(* IEC 61131-3 sources: iecf/harness/cases (part 5) *)

(* ---- narrowingcompare.st ---- *)
(* implicit-narrowing: a ULINT and a signed integer, which no type holds
   both of, compared by their values, W0010 at each - as TcOpen's tests'
   `_plcCycleCounter >= _reqStep + 7`, a ULINT and an INT. Worked by
   hand, u 5, m -1, big 2^64 - 1, l -1, seven 7, four 4:
   u > m TRUE (%QX0.0); m < u TRUE (%QX0.1); u = m FALSE (%QX0.2);
   big > l TRUE, where the bits alike would say equal (%QX0.3);
   u + 2 = seven, 7 = 7, TRUE (%QX0.4); u <= four FALSE (%QX0.5).
   reference-skip: implicit narrowing is CODESYS's, not IEC 61131-3. *)
PROGRAM main
  VAR
    u : ULINT := 5; big : ULINT := 18446744073709551615;
    m : INT := -1; l : LINT := -1; seven : DINT := 7; four : SINT := 4;
  END_VAR
  VAR
    q0 AT %QX0.0 : BOOL; q1 AT %QX0.1 : BOOL; q2 AT %QX0.2 : BOOL;
    q3 AT %QX0.3 : BOOL; q4 AT %QX0.4 : BOOL; q5 AT %QX0.5 : BOOL;
  END_VAR
  q0 := u > m;
  q1 := m < u;
  q2 := u = m;
  q3 := big > l;
  q4 := u + 2 = seven;
  q5 := u <= four;
END_PROGRAM

CONFIGURATION cf
  RESOURCE r ON x
    TASK tk(INTERVAL := T#10ms, PRIORITY := 1);
    PROGRAM p WITH tk : main;
  END_RESOURCE
END_CONFIGURATION

(* ---- narrowingliteral.st ---- *)
(* implicit-narrowing: an integer literal outside the integer or bit
   string type it goes into keeps its low bits, as a conversion of a
   typed one would, W0010 at each - as TcOpen's `_testId := -1` of a
   ULINT and `_theOrderOfThePreviouslyExecutedStep := -1` of a UINT.
   Worked by hand:
   u := -1, a UINT: 65535, 16#FFFF (%QW0).
   g(300), to a USINT input: 300 - 256, 44, 16#2C (%QB2).
   s := 200, a SINT: 200 - 256, -56, 16#C8 (%QB3).
   w := 16#12345, a WORD: 16#2345 (%QW4).
   l := -1, a ULINT: 2^64 - 1, all ones (%QL8).
   i, initialised to -2, a UDINT: 2^32 - 2, 16#FFFFFFFE (%QD16).
   reference-skip: implicit narrowing is CODESYS's, not IEC 61131-3. *)
FUNCTION g : USINT
  VAR_INPUT x : USINT; END_VAR
  g := x;
END_FUNCTION

PROGRAM main
  VAR
    u : UINT; s : SINT; w : WORD; l : ULINT; i : UDINT := -2;
  END_VAR
  VAR
    q0 AT %QW0 : UINT; q1 AT %QB2 : USINT; q2 AT %QB3 : SINT; q3 AT %QW4 : WORD;
    q4 AT %QL8 : ULINT; q5 AT %QD16 : UDINT;
  END_VAR
  u := -1;
  q0 := u;
  q1 := g(300);
  s := 200;
  q2 := s;
  w := 16#12345;
  q3 := w;
  l := -1;
  q4 := l;
  q5 := i;
END_PROGRAM

CONFIGURATION cf
  RESOURCE r ON x
    TASK tk(INTERVAL := T#10ms, PRIORITY := 1);
    PROGRAM p WITH tk : main;
  END_RESOURCE
END_CONFIGURATION

(* ---- narrowingreal.st ---- *)
(* implicit-narrowing: an integer where a real is wanted and Figure 11
   has no implicit conversion, and an LREAL where a REAL is, converted
   as DINT_TO_REAL and LREAL_TO_REAL would, W0010 at each - as TcOpen's
   `_price := Price` (an LREAL property into a REAL), its
   TcoBytesToReal's LREAL into the REAL result, and a DINT given to
   TcoRealToBytes's `inValue : REAL`. Worked by hand:
   r := d, DINT 16777217 into a REAL: the nearest REAL, 16777216.0,
   16#4B800000 (%QD0).
   r := l, LREAL 1.5: 1.5, 16#3FC00000 (%QD4).
   twice(n), the DINT 3 to a REAL input: 6.0, 16#40C00000 (%QD8).
   quarter(), an LREAL 2.25 into the REAL result: 16#40100000 (%QD12).
   reference-skip: implicit narrowing is CODESYS's, not IEC 61131-3. *)
FUNCTION twice : REAL
  VAR_INPUT x : REAL; END_VAR
  twice := x * 2.0;
END_FUNCTION

FUNCTION quarter : REAL
  VAR l : LREAL := 2.25; END_VAR
  quarter := l;
END_FUNCTION

PROGRAM main
  VAR
    d : DINT := 16777217; l : LREAL := 1.5; n : DINT := 3; r : REAL;
  END_VAR
  VAR
    q0 AT %QD0 : REAL;
    q1 AT %QD4 : REAL;
    q2 AT %QD8 : REAL;
    q3 AT %QD12 : REAL;
  END_VAR
  r := d;
  q0 := r;
  r := l;
  q1 := r;
  q2 := twice(n);
  q3 := quarter();
END_PROGRAM

CONFIGURATION cf
  RESOURCE r ON x
    TASK tk(INTERVAL := T#10ms, PRIORITY := 1);
    PROGRAM p WITH tk : main;
  END_RESOURCE
END_CONFIGURATION

(* ---- nesten.st ---- *)
(* Calls with EN nested in another's arguments, and EN on a FUNCTION
   giving an array or a structure (Ed.3 6.6.1.5; docs/dependencies.md:
   EN FALSE does not evaluate the inputs, calls nothing and leaves the
   statement undone). Worked by hand:
   b TRUE: ADD(EN := b, IN1 := ADD(EN := b, IN1 := 1, IN2 := 2),
   IN2 := 3): 6 (%QB0). b FALSE, v 9 before: the statement is undone, v
   9 (%QB1).
   t 32767: ADD(EN := TRUE, IN1 := ADD(EN := TRUE, IN1 := t, IN2 := 1,
   ENO => e2), IN2 := 0, ENO => e1): the inner one overflows, wraps to
   -32768 and is flagged OVERFLOW, its ENO FALSE (%QX2.0 0); the outer
   adds 0, no flag of its own: its ENO TRUE (%QX2.1 1); v / 1000 is -32
   (%QB3).
   Inc adds 1 to its in-out. n 0: ADD(EN := TRUE, IN1 := Inc(EN :=
   TRUE, io := n), IN2 := 10): 11 (%QB4), n 1 (%QB5). The outer's EN
   FALSE, v 5 before: Inc is not called, v 5 (%QB6), n still 1 (%QB7).
   FA gives [x, 2x, 0]: a := FA(EN := TRUE, x := 4), a[2] 8 (%QB8);
   a := FA(EN := FALSE, x := 7) leaves a: a[1] 4 (%QB9).
   p := FP(EN := TRUE, x := 3, ENO => e3): p.x 3 (%QB10), e3 TRUE
   (%QX11.0). SumA(FA(EN := TRUE, x := 2)), 2 + 4 + 0: 6 (%QB12).
   The first flag is the inner ADD's OVERFLOW.
   reference-skip: a nested call with ENO or an in-out, an array
   input: its C does not build. *)
TYPE
  A3 : ARRAY [1..3] OF INT;
  PT : STRUCT x : INT; END_STRUCT;
END_TYPE
FUNCTION Inc : INT
  VAR_IN_OUT io : INT; END_VAR
  io := io + 1;
  Inc := io;
END_FUNCTION
FUNCTION FA : A3
  VAR_INPUT x : INT; END_VAR
  FA[1] := x;
  FA[2] := x * 2;
END_FUNCTION
FUNCTION FP : PT
  VAR_INPUT x : INT; END_VAR
  FP.x := x;
END_FUNCTION
FUNCTION SumA : INT
  VAR_INPUT q : A3; END_VAR
  SumA := q[1] + q[2] + q[3];
END_FUNCTION
PROGRAM main
  VAR
    b : BOOL := TRUE;
    v : INT;
    t : INT := 32767;
    n : INT;
    e1 : BOOL;
    e2 : BOOL;
    e3 : BOOL;
    a : A3;
    p : PT;
  END_VAR
  VAR
    q0 AT %QB0 : SINT;
    q1 AT %QB1 : SINT;
    q20 AT %QX2.0 : BOOL;
    q21 AT %QX2.1 : BOOL;
    q3 AT %QB3 : SINT;
    q4 AT %QB4 : SINT;
    q5 AT %QB5 : SINT;
    q6 AT %QB6 : SINT;
    q7 AT %QB7 : SINT;
    q8 AT %QB8 : SINT;
    q9 AT %QB9 : SINT;
    q10 AT %QB10 : SINT;
    q11 AT %QX11.0 : BOOL;
    q12 AT %QB12 : SINT;
  END_VAR
  v := ADD(EN := b, IN1 := ADD(EN := b, IN1 := 1, IN2 := 2), IN2 := 3);
  q0 := INT_TO_SINT(v);
  b := FALSE;
  v := 9;
  v := ADD(EN := b, IN1 := ADD(EN := b, IN1 := 1, IN2 := 2), IN2 := 3);
  q1 := INT_TO_SINT(v);
  v := ADD(EN := TRUE, IN1 := ADD(EN := TRUE, IN1 := t, IN2 := 1, ENO => e2), IN2 := 0, ENO => e1);
  q20 := e2;
  q21 := e1;
  q3 := INT_TO_SINT(v / 1000);
  n := 0;
  v := ADD(EN := TRUE, IN1 := Inc(EN := TRUE, io := n), IN2 := 10);
  q4 := INT_TO_SINT(v);
  q5 := INT_TO_SINT(n);
  v := 5;
  v := ADD(EN := FALSE, IN1 := Inc(EN := TRUE, io := n), IN2 := 10);
  q6 := INT_TO_SINT(v);
  q7 := INT_TO_SINT(n);
  a := FA(EN := TRUE, x := 4);
  q8 := INT_TO_SINT(a[2]);
  a := FA(EN := FALSE, x := 7);
  q9 := INT_TO_SINT(a[1]);
  p := FP(EN := TRUE, x := 3, ENO => e3);
  q10 := INT_TO_SINT(p.x);
  q11 := e3;
  q12 := INT_TO_SINT(SumA(FA(EN := TRUE, x := 2)));
END_PROGRAM

CONFIGURATION c
  RESOURCE r ON x
    TASK t(INTERVAL := T#10ms, PRIORITY := 1);
    PROGRAM p WITH t : main;
  END_RESOURCE
END_CONFIGURATION

(* ---- overflow.st ---- *)
(* Where iecf differs from the reference compiler on purpose (PROPOSAL.md §6.3): an
   integer overflow is flagged. At tick 2, a + b leaves INT. Both wrap to
   -1536 and go on, as CODESYS, TwinCAT, Siemens and Rockwell do; iecf
   also records the first overflow, its POU and line, in ctx->flag, which
   stays until the platform clears it. Its trace is overflow.iecf.trace:
   the reference compiler's bytes, with "flag 2 MAIN 18" from tick 2.

   MOD by zero is 0 in both: Ed.3 Table 29 e defines it so. *)
PROGRAM main
VAR
  a AT %IW0 : INT;
  b AT %IW2 : INT;
  r_mod AT %MW0 : INT;
  r_sum AT %MW2 : INT;
  after AT %MW4 : INT;
END_VAR
r_mod := a MOD b;
r_sum := a + b;
after := after + 1;
END_PROGRAM

CONFIGURATION plant
  RESOURCE r ON PLC
    TASK fast(INTERVAL := T#10ms, PRIORITY := 0);
    PROGRAM p WITH fast : main;
  END_RESOURCE
END_CONFIGURATION

(* ---- parts.st ---- *)
(* CONCAT_DATE, CONCAT_TOD, CONCAT_DT and the SPLITs (Ed.3 Table 36;
   docs/dependencies.md): a month from 11 and an hour from 22 go up by one
   each tick, joined into a DATE, a TOD and a DT and split back. The parts
   are valid at tick 1 (2026-12-31, 23:30:15.250); a day not in its month
   (November 31st, at tick 0), a month 13 or an hour 24 gives the type's
   default value in iecf, flagged; iecf's trace is parts.iecf.trace. *)
PROGRAM main
VAR
  r_year AT %MW0 : UINT;
  r_month AT %MB2 : USINT;
  r_day AT %MB3 : USINT;
  r_hour AT %MB4 : USINT;
  r_min AT %MB5 : USINT;
  r_sec AT %MB6 : USINT;
  r_ms AT %MW8 : UINT;
  r_dt_month AT %MB10 : USINT;
  r_dt_hour AT %MB11 : USINT;
END_VAR
VAR
  month : INT := 10;
  hour : SINT := 21;
  d : DATE;
  t : TOD;
  s : DT;
  y, m, dd : UDINT;
END_VAR
month := month + 1;
hour := hour + 1;
d := CONCAT_DATE(2026, month, 31);
t := CONCAT_TOD(hour, 30, 15, 250);
s := CONCAT_DT(YEAR := 2026, MONTH := month, DAY := 28, HOUR := hour,
               MINUTE := 59, SECOND := 59, MILLISECOND := 999);
SPLIT_DATE(d, y, m, dd);
r_year := UDINT_TO_UINT(y);
r_month := UDINT_TO_USINT(m);
r_day := UDINT_TO_USINT(dd);
SPLIT_TOD(IN := t, HOUR => r_hour, MINUTE => r_min, SECOND => r_sec, MILLISECOND => r_ms);
SPLIT_DT(IN := s, MONTH => r_dt_month, HOUR => r_dt_hour);
END_PROGRAM

CONFIGURATION plant
  RESOURCE r ON PLC
    TASK fast(INTERVAL := T#10ms, PRIORITY := 0);
    PROGRAM p WITH fast : main;
  END_RESOURCE
END_CONFIGURATION

(* ---- pointerfault.st ---- *)
(* A pointer read past its variable (the pointers extension): a fault,
   IECF_FAULT_INDEX, the task stopped where the read leaves the variable,
   never C's undefined behaviour. Worked by hand: a has 4 bytes, 1 2 3 4;
   the loop adds them through pt for i 0..4, so the fifth read, past the
   end, faults on line 21 in the first tick, n holding 10 so far, and
   the task stops there: %QB0, set after the loop, stays 0. (The host
   leaves the fault set, so a later tick stops at once: whether to run
   again is the platform's; %QB1 is the first statement's, 0.)
   reference-skip: pointers are CODESYS's, not IEC 61131-3. *)
PROGRAM main
  VAR
    a : ARRAY[0..3] OF BYTE := [1, 2, 3, 4];
    pt : POINTER TO BYTE;
    i, n : INT;
  END_VAR
  VAR q0 AT %QB0 : SINT; q1 AT %QB1 : SINT; END_VAR
  q1 := INT_TO_SINT(n);
  n := 0;
  pt := ADR(a);
  FOR i := 0 TO 4 DO
    n := n + BYTE_TO_INT(pt^);
    pt := pt + 1;
  END_FOR;
  q0 := INT_TO_SINT(n);
END_PROGRAM

CONFIGURATION cf
  RESOURCE r ON x
    TASK tk(INTERVAL := T#10ms, PRIORITY := 1);
    PROGRAM p WITH tk : main;
  END_RESOURCE
END_CONFIGURATION

(* ---- pointerindex.st ---- *)
(* A pointer indexed (the pointers extension): p[i] is (p + i *
   SIZEOF(T))^, as CODESYS and TwinCAT index a pointer, checked as p^
   is. Worked by hand: a is 10 20 30 40 50, so the loop adds 150 and
   %QB0 is 15; p[k] with k 2 writes a[2] := 7; p moved to ADR(p[3]),
   a[3], reads p[-1] + p[0], 7 + 40, so %QB1 is 47; q[1].y := 9 and
   s[2].x := 4 read back through q and s, 9 + 4, %QB2 13; p[1] is
   a[4], 50, %QB3 5; %QB4 set to 1, then p[2] is past a's end: a
   fault, IECF_FAULT_INDEX, on line 36, %QB4 left at 1.
   reference-skip: pointers are CODESYS's, not IEC 61131-3. *)
TYPE pair : STRUCT x : INT; y : INT; END_STRUCT; END_TYPE
PROGRAM main
  VAR
    a : ARRAY[0..4] OF INT := [10, 20, 30, 40, 50];
    s : ARRAY[0..2] OF pair;
    p : POINTER TO INT;
    q : POINTER TO pair;
    i, n : INT;
    k : UINT := 2;
  END_VAR
  VAR q0 AT %QB0 : SINT; q1 AT %QB1 : SINT; q2 AT %QB2 : SINT; q3 AT %QB3 : SINT; q4 AT %QB4 : SINT; END_VAR
  p := ADR(a);
  n := 0;
  FOR i := 0 TO 4 DO
    n := n + p[i];
  END_FOR;
  q0 := INT_TO_SINT(n / 10);
  p[k] := 7;
  p := ADR(p[3]);
  q1 := INT_TO_SINT(p[-1] + p[0]);
  q := ADR(s);
  q[1].y := 9;
  s[2].x := 4;
  q2 := INT_TO_SINT(s[1].y + q[2].x);
  q3 := INT_TO_SINT(p[1] / 10);
  q4 := 1;
  q4 := INT_TO_SINT(p[2]);
END_PROGRAM

CONFIGURATION cf
  RESOURCE r ON x
    TASK tk(INTERVAL := T#10ms, PRIORITY := 1);
    PROGRAM p WITH tk : main;
  END_RESOURCE
END_CONFIGURATION

(* ---- pointers.st ---- *)
(* Pointers (the pointers extension), in the ways the OSCAT BASIC library
   uses them. Worked by hand:
   %QB0: StrLen walks a STRING's bytes through a POINTER TO BYTE to its
   0: 'hello', 5.
   %QB1: Sum takes ADR(a) and SIZEOF(a) of an ARRAY[0..3] OF REAL, as
   OSCAT's array functions do, and counts SIZEOF(a) / SIZEOF(pt^[0]) = 4
   elements: 1.5 + 2.5 + 3.0 + 4.0 = 11.0, as SINT 11.
   %QB2: Clear zeroes a BYTE buffer by pointer arithmetic, pt < stop,
   pt := pt + 1, from ADR(buf) to ADR(buf) + SIZEOF(buf); then buf[0] +
   buf[7], 0.
   %QB3: four bytes 16#11 16#22 16#33 16#44 read as one DWORD through a
   POINTER TO DWORD: 16#44332211 on a little-endian platform, its low
   byte 16#11.
   %QB4: a structure's field through a pointer, s.b := 7 by ps^.b := 7;
   and ps^.a + ps^.b with a 2: 9.
   %QB5: two pointers into one array subtracted: ADR(a[3]) - ADR(a[0]),
   3 * SIZEOF(REAL), 12.
   reference-skip: pointers are CODESYS's, not IEC 61131-3. *)
TYPE Pair : STRUCT a : SINT; b : SINT; END_STRUCT; END_TYPE

FUNCTION StrLen : INT
  VAR_INPUT pt : POINTER TO BYTE; END_VAR
  StrLen := 0;
  WHILE pt^ <> 0 DO
    StrLen := StrLen + 1;
    pt := pt + 1;
  END_WHILE;
END_FUNCTION

FUNCTION Sum : REAL
  VAR_INPUT pt : POINTER TO ARRAY[0..32000] OF REAL; size : UINT; END_VAR
  VAR i : INT; END_VAR
  Sum := 0.0;
  FOR i := 0 TO UINT_TO_INT(size / SIZEOF(pt^[0])) - 1 DO
    Sum := Sum + pt^[i];
  END_FOR;
END_FUNCTION

FUNCTION Clear : BOOL
  VAR_INPUT pt : POINTER TO BYTE; size : UINT; END_VAR
  VAR stop : POINTER TO BYTE; END_VAR
  stop := pt + size;
  WHILE pt < stop DO
    pt^ := 0;
    pt := pt + 1;
  END_WHILE;
  Clear := TRUE;
END_FUNCTION

PROGRAM main
  VAR
    s : STRING[20] := 'hello';
    a : ARRAY[0..3] OF REAL := [1.5, 2.5, 3.0, 4.0];
    buf : ARRAY[0..7] OF BYTE := [8(16#FF)];
    bytes : ARRAY[0..3] OF BYTE := [16#11, 16#22, 16#33, 16#44];
    pd : POINTER TO DWORD;
    pr : Pair := (a := 2);
    ps : POINTER TO Pair;
    ok : BOOL;
  END_VAR
  VAR
    q0 AT %QB0 : SINT; q1 AT %QB1 : SINT; q2 AT %QB2 : BYTE; q3 AT %QB3 : BYTE;
    q4 AT %QB4 : SINT; q5 AT %QB5 : SINT;
  END_VAR
  q0 := INT_TO_SINT(StrLen(ADR(s)));
  q1 := REAL_TO_SINT(Sum(ADR(a), SIZEOF(a)));
  ok := Clear(ADR(buf), SIZEOF(buf));
  q2 := buf[0] OR buf[7];
  pd := ADR(bytes);
  q3 := DWORD_TO_BYTE(pd^);
  ps := ADR(pr);
  ps^.b := 7;
  q4 := ps^.a + ps^.b;
  q5 := DINT_TO_SINT(ADR(a[3]) - ADR(a[0]));
END_PROGRAM

CONFIGURATION cf
  RESOURCE r ON x
    TASK tk(INTERVAL := T#10ms, PRIORITY := 1);
    PROGRAM p WITH tk : main;
  END_RESOURCE
END_CONFIGURATION

(* ---- pointers2.st ---- *)
(* Pointers (the pointers extension): a STRING whole through a pointer,
   arrays and structures copied whole through one, ADR of a variable at
   an address, and ADR() as an initial value. Worked by hand:
   %QB0: ps := ADR(s); ps^ := 'abc' writes the STRING through ps; then
   LEN(s), 3.
   %QB1: t := ps^ reads it back whole; LEN(t) + LEN(ps^), 3 + 3 = 6.
   %QB2: pa := ADR(src); dst := pa^ copies the array [5, 6, 7] whole;
   dst[2], 7.
   %QB3: pq^ := pr copies a structure whole into r2 (pq := ADR(r2)), then
   r2.b, 9.
   %QB4: pin points at %IB2, ADR of a variable at an address; the
   input bytes are 0, so pin^ reads 0; pq0 points at the output %QB5 and
   writes 16#2A through it (%QB5), read back as 42 into %QB4.
   %QB6: pinit's initial value ADR(src[1]) points at src[1], 6.
   reference-skip: pointers are CODESYS's, not IEC 61131-3. *)
TYPE R : STRUCT a : SINT; b : SINT; END_STRUCT; END_TYPE

PROGRAM main
  VAR
    s : STRING[20];
    t : STRING[20];
    ps : POINTER TO STRING[20];
    src : ARRAY[0..2] OF SINT := [5, 6, 7];
    dst : ARRAY[0..2] OF SINT;
    pa : POINTER TO ARRAY[0..2] OF SINT;
    pr : R := (a := 1, b := 9);
    r2 : R;
    pq : POINTER TO R;
    pinit : POINTER TO SINT := ADR(src[1]);
    pin : POINTER TO BYTE;
    pq0 : POINTER TO BYTE;
  END_VAR
  VAR
    q0 AT %QB0 : SINT; q1 AT %QB1 : SINT; q2 AT %QB2 : SINT; q3 AT %QB3 : SINT;
    q4 AT %QB4 : BYTE; q5 AT %QB5 : BYTE; q6 AT %QB6 : SINT;
    i2 AT %IB2 : BYTE;
  END_VAR
  ps := ADR(s);
  ps^ := 'abc';
  q0 := INT_TO_SINT(LEN(s));
  t := ps^;
  q1 := INT_TO_SINT(LEN(t) + LEN(ps^));
  pa := ADR(src);
  dst := pa^;
  q2 := dst[2];
  pq := ADR(r2);
  pq^ := pr;
  q3 := r2.b;
  pin := ADR(i2);
  pq0 := ADR(q5);
  pq0^ := pin^ + 16#2A;
  q4 := q5;
  q6 := pinit^;
END_PROGRAM

CONFIGURATION cf
  RESOURCE r ON x
    TASK tk(INTERVAL := T#10ms, PRIORITY := 1);
    PROGRAM p WITH tk : main;
  END_RESOURCE
END_CONFIGURATION

(* ---- progio.st ---- *)
(* A program's VAR_IN_OUT (Ed.3 Table 47 2c), connected in the
   CONFIGURATION to a global (6.8.2): each instance of `bump` reads and
   writes the global itself, through its in-out. Two instances on one
   task add 1 and 10 to `shared` each tick, a third program copies it to
   %MW0; `other` is never touched. The reference compiler cannot compile
   program connections (PROPOSAL.md §1b): iecf only, a hand-checked
   trace. *)
PROGRAM bump
VAR_INPUT amount : INT; END_VAR
VAR_IN_OUT n : INT; END_VAR
n := n + amount;
END_PROGRAM

PROGRAM show
VAR_EXTERNAL shared, other : INT; END_VAR
VAR
  r_shared AT %MW0 : INT;
  r_other AT %MW2 : INT;
END_VAR
r_shared := shared;
r_other := other;
END_PROGRAM

CONFIGURATION plant
  VAR_GLOBAL shared : INT := 100; other : INT := 7; END_VAR
  RESOURCE r ON PLC
    TASK fast(INTERVAL := T#10ms, PRIORITY := 0);
    PROGRAM one WITH fast : bump(amount := 1, n := shared);
    PROGRAM ten WITH fast : bump(amount := 10, n := shared);
    PROGRAM s WITH fast : show;
  END_RESOURCE
END_CONFIGURATION

(* ---- real.st ---- *)
(* REAL and LREAL: arithmetic, comparisons, conversions to and from the
   integers, and the functions of Ed.3 Table 28 whose results are exact in
   binary floating point. REAL_TO_INT rounds halves to even, as Ed.3
   Table 22's examples have it (2.5 to 2, -2.5 to -2).

   Truncation is the deprecated TRUNC (Ed.3 Table 22 2a; W0003 in iecf),
   the one form the reference compiler also knows, into a DINT: the reference compiler types it by its
   target, iecf gives DINT as the vendors do (docs/dependencies.md). *)
PROGRAM main
VAR
  inp AT %IW0 : INT;
  r_add AT %MD0 : REAL;
  r_mul AT %MD4 : REAL;
  r_div AT %ML8 : LREAL;
  r_round AT %MW16 : INT;
  r_trunc AT %MD38 : DINT;
  r_sqrt AT %MD20 : REAL;
  r_abs AT %ML24 : LREAL;
  r_cmp AT %MB32 : BYTE;
  r_lr AT %MD34 : REAL;
END_VAR
VAR
  x : REAL;
  y : LREAL;
END_VAR
x := INT_TO_REAL(inp) / 4.0;
y := INT_TO_LREAL(inp) * 0.5;
r_add := x + 1.5;
r_mul := x * -2.0;
r_div := y / 3.0;
r_round := REAL_TO_INT(x);
r_trunc := TRUNC(x);
r_sqrt := SQRT(ABS(x) * ABS(x));
r_abs := ABS(y - 100.0);
r_cmp := 0;
IF x > 1.0 THEN r_cmp := r_cmp OR 1; END_IF;
IF y <= -1.0 THEN r_cmp := r_cmp OR 2; END_IF;
IF x = 2.5 THEN r_cmp := r_cmp OR 4; END_IF;
r_lr := LREAL_TO_REAL(y) + 0.25;
END_PROGRAM

CONFIGURATION plant
  RESOURCE r ON PLC
    TASK fast(INTERVAL := T#10ms, PRIORITY := 0);
    PROGRAM p WITH fast : main;
  END_RESOURCE
END_CONFIGURATION

(* ---- realchains.st ---- *)
(* REAL and LREAL chains tested once (docs/c-output.md §5, chains.rs),
   through a standard function, a conversion, an array element and a
   divisor that is itself a result: an infinity or NaN at each, one a
   tick, the flag cleared before each (`unflag`), flagged as each
   operator tested on its own flags it - by its code and line. The
   trace is the one iecf gave before chains took these in.
   tick 0 the set-up's overflow at line 26 (x * x), the rest finite.
   tick 1 SIN of an overflowing product: overflow (flag 2), line 30.
   tick 2 LN(0.0) plus one: -infinity, overflow, line 31.
   tick 3 SQRT(-1.0) times two: NaN (flag 9), line 32.
   tick 4 EXP of minus an infinite input: 0, nothing flagged.
   tick 5 LREAL_TO_REAL(1.0E300) plus one: overflow, line 34.
   tick 6 an infinite array element times 2 plus 1: overflow, line 35.
   tick 7 divided by an overflowing product: overflow, line 36; the
          quotient 0, %QD0 2000.
   tick 8 ABS and ATAN of a leaf, COS, TAN, ASIN(2.0): NaN, line 37.
   tick 9 DINT_TO_LREAL(i) times 1.0E308 times 10: overflow, line 38.
   tick 10 divided by a difference of 0: the fault, line 39; no tick
          runs after it.
   %QD0 a finite witness, %QB4 the tick.
   reference-skip: its own flags; the reference compiler has none. *)
PROGRAM main
  VAR k : USINT; x : LREAL := 1.0E200; y : LREAL; inf : LREAL; i : DINT := 7;
      r : REAL; a : ARRAY[1..3] OF LREAL; n : INT := 2; zero : LREAL; w : LREAL; END_VAR
  VAR q0 AT %QD0 : DINT; q1 AT %QB4 : USINT; END_VAR
  IF k = 0 THEN inf := x * x; END_IF;
  IF k = 0 THEN a[n] := x * x; END_IF;
  CASE k OF
    0: y := SIN(0.5) * COS(0.5) + SQRT(4.0) / (1.0 + 2.0 * 3.0); w := y;
    1: y := SIN(x * x) + 1.0;
    2: y := LN(zero) + 1.0;
    3: y := SQRT(-1.0) * 2.0;
    4: y := EXP(-inf) * 2.0 + 1.0; w := y;
    5: r := LREAL_TO_REAL(1.0E300) + 1.0;
    6: y := a[n] * 2.0 + 1.0;
    7: y := 1.0 / (x * x) + 2.0; w := y;
    8: y := ABS(-x) * 0.0 + ATAN(2.0) + COS(0.1) * TAN(0.2) + ASIN(2.0);
    9: y := DINT_TO_LREAL(i) * 1.0E308 * 10.0;
    10: y := 1.0 / (x - x) + 2.0;
  END_CASE;
  q0 := LREAL_TO_DINT(w * 1000.0);
  q1 := k;
  k := k + 1;
END_PROGRAM
CONFIGURATION cf
  RESOURCE r ON x
    TASK tk(INTERVAL := T#10ms, PRIORITY := 1);
    PROGRAM p WITH tk : main;
  END_RESOURCE
END_CONFIGURATION

(* ---- refgated.st ---- *)
(* REF() of an element whose index is a call with EN and ENO: the call
   made once, its ENO taken. Worked by hand: the index is ADD(1, 2), 3,
   so r refers to a[3], 30 (Q0 1e); ENO TRUE (Q1 01).
   The same on the reference compiler. *)
PROGRAM main
  VAR a : ARRAY [1..4] OF INT := [10, 20, 30, 40]; r : REF_TO INT; b : BOOL := TRUE; ok : BOOL; END_VAR
  VAR q AT %QB0 : USINT; q1 AT %QB1 : USINT; END_VAR
  r := REF(a[ADD(EN := b, IN1 := 1, IN2 := 2, ENO => ok)]);
  q := INT_TO_USINT(r^);
  q1 := BOOL_TO_USINT(ok);
END_PROGRAM
CONFIGURATION c RESOURCE r ON PLC TASK t(INTERVAL := T#10ms, PRIORITY := 1); PROGRAM p WITH t : main; END_RESOURCE END_CONFIGURATION

(* ---- resaccess.st ---- *)
(* A global named through its resource (Ed.3 6.8.2, Global_Var_Access):
   `R.g` and `R.g.x` in a program's connections - an input, an output,
   an in-out - and in a TASK's INTERVAL, beside the plain names. r1's
   task runs every 20 ms, on ticks 0 and 2; r2's every tick, after it.
   Worked by hand:

   tick 0, r1.m: a 10, b p.y 4: o 14 into res (Q0 0e 00), o2 6 into
   p.x, cnt 1. r1.w: a p.x 6, b cnt 1: o 7 (Q2 07 00); its in-out is the
   configuration's g, 2. r2.m: a its own g1 20, b g 2: o 22 (Q4 16 00),
   o2 18 (Q6 12 00).
   tick 1: r2.m alone, the same.
   tick 2, r1.m: 14, 6, cnt 2. r1.w: 6 + 2 = 8 (08 00), g 3. r2.m: 20 +
   3 = 23 (17 00), 17 (11 00).
   reference-skip: program connections, as `connections`. *)
TYPE Pt : STRUCT x : INT; y : INT; END_STRUCT; END_TYPE
PROGRAM main
  VAR_INPUT a : INT; b : INT; END_VAR
  VAR_OUTPUT o : INT; o2 : INT; END_VAR
  VAR_IN_OUT n : INT; END_VAR
  o := a + b;
  o2 := a - b;
  n := n + 1;
END_PROGRAM
CONFIGURATION plant
  VAR_GLOBAL g : INT := 1; END_VAR
  RESOURCE r1 ON PLC
    VAR_GLOBAL g1 : INT := 10; p : Pt := (x := 3, y := 4); cnt : INT; iv : TIME := T#20ms; END_VAR
    VAR_GLOBAL res AT %QW0 : INT; res2 AT %QW2 : INT; END_VAR
    TASK t(INTERVAL := r1.iv, PRIORITY := 1);
    PROGRAM m WITH t : main(a := r1.g1, b := r1.p.y, o => r1.res, o2 => r1.p.x, n := r1.cnt);
    PROGRAM w WITH t : main(a := r1.p.x, b := r1.cnt, o => res2, n := g);
  END_RESOURCE
  RESOURCE r2 ON PLC
    VAR_GLOBAL g1 : INT := 20; cnt : INT; END_VAR
    VAR_GLOBAL res AT %QW4 : INT; out2 AT %QW6 : INT; END_VAR
    TASK t(INTERVAL := T#10ms, PRIORITY := 2);
    PROGRAM m WITH t : main(a := r2.g1, b := g, o => r2.res, o2 => out2, n := r2.cnt);
  END_RESOURCE
END_CONFIGURATION

(* ---- retain.st ---- *)
(* RETAIN (Ed.3 6.5.6): a warm restart sets every variable to its initial
   value but the RETAIN ones, which keep theirs (docs/c-output.md §7); a
   cold start sets them too. Globals and a program's variables, a whole
   function block instance among them, count each tick. At tick 3 a warm
   restart: the plain counters start again, the RETAIN ones go on.
   The reference compiler has no warm restart of its own; its host starts everything
   anew. iecf's trace is retain.iecf.trace. *)
PROGRAM main
VAR_EXTERNAL
  g_plain : INT;
  g_kept : INT;
END_VAR
VAR
  r_plain AT %MW0 : INT;
  r_kept AT %MW2 : INT;
  r_g_plain AT %MW4 : INT;
  r_g_kept AT %MW6 : INT;
  r_ctu AT %MW8 : INT;
  r_arr AT %MW10 : INT;
END_VAR
VAR
  plain : INT := 100;
END_VAR
VAR RETAIN
  kept : INT := 100;
  c : CTU;
  arr : ARRAY [1..2] OF INT := [7, 8];
END_VAR
plain := plain + 1;
kept := kept + 1;
g_plain := g_plain + 1;
g_kept := g_kept + 1;
c(CU := NOT c.CU, PV := 1000);
arr[2] := arr[2] + 1;
r_plain := plain;
r_kept := kept;
r_g_plain := g_plain;
r_g_kept := g_kept;
r_ctu := c.CV;
r_arr := arr[2];
END_PROGRAM

CONFIGURATION plant
  VAR_GLOBAL g_plain : INT; END_VAR
  VAR_GLOBAL RETAIN g_kept : INT := 50; END_VAR
  RESOURCE r ON PLC
    TASK fast(INTERVAL := T#10ms, PRIORITY := 0);
    PROGRAM p WITH fast : main;
  END_RESOURCE
END_CONFIGURATION

(* ---- sfc.st ---- *)
(* SFC (Ed.3 6.7; docs/behaviour/sfc.md): one scan runs the action
   control, the actions (those ending first), then the transitions of the
   steps active when it began. S1 holds every kind of association: a BOOL
   variable as an action (lamp, N), S and R (Sto, reset in S4), L and D of
   20 ms (Lim, Del), P1 and P0 (Ent, Ext); its transition waits for
   S1.T >= T#40ms, then divides into S2 and S3, which converge into S4.
   From S4 two transitions: (PRIORITY := 1) back to S0 when back, else
   (PRIORITY := 2) to S5. Ent RETURNs after counting: only the action
   ends. The x outputs show the active steps (BOOL variables as N
   actions). A scan is 10 ms. The reference compiler tests transitions first and has no
   final scan, nor PRIORITY: this case is iecf's alone (reference-skip),
   its trace checked by hand. *)
PROGRAM main
VAR
  go AT %IX0.0 : BOOL;
  back AT %IX0.1 : BOOL;
  lamp AT %QX0.0 : BOOL;
  stored AT %QX0.1 : BOOL;
  limited AT %QX0.2 : BOOL;
  delayed AT %QX0.3 : BOOL;
  nent AT %QB1 : USINT;
  next AT %QB2 : USINT;
  x0 AT %QX3.0 : BOOL;
  x1 AT %QX3.1 : BOOL;
  x2 AT %QX3.2 : BOOL;
  x3 AT %QX3.3 : BOOL;
  x4 AT %QX3.4 : BOOL;
  x5 AT %QX3.5 : BOOL;
END_VAR

INITIAL_STEP S0:
  x0(N);
END_STEP
STEP S1:
  x1(N);
  lamp(N);
  Sto(S);
  Lim(L, T#20ms);
  Del(D, T#20ms);
  Ent(P1);
  Ext(P0);
END_STEP
STEP S2:
  x2(N);
END_STEP
STEP S2b:
END_STEP
STEP S3:
  x3(N);
END_STEP
STEP S4:
  x4(N);
  Sto(R);
END_STEP
STEP S5:
  x5(N);
END_STEP

TRANSITION FROM S0 TO S1 := go; END_TRANSITION
TRANSITION FROM S1 TO (S2, S3) := S1.T >= T#40ms; END_TRANSITION
TRANSITION FROM S2 TO S2b := TRUE; END_TRANSITION
TRANSITION FROM (S2b, S3) TO S4 := TRUE; END_TRANSITION
TRANSITION (PRIORITY := 2) FROM S4 TO S5 := TRUE; END_TRANSITION
TRANSITION (PRIORITY := 1) FROM S4 TO S0 := back; END_TRANSITION
TRANSITION FROM S5 TO S0 := TRUE; END_TRANSITION

ACTION Sto:
  stored := Sto.Q;
END_ACTION
ACTION Lim:
  limited := Lim.Q;
END_ACTION
ACTION Del:
  delayed := Del.Q;
END_ACTION
ACTION Ent:
  nent := nent + 1;
  RETURN;
  nent := nent + 100;
END_ACTION
ACTION Ext:
  next := next + 1;
END_ACTION
END_PROGRAM

CONFIGURATION plant
  RESOURCE res ON PLC
    TASK fast(INTERVAL := T#10ms, PRIORITY := 0);
    PROGRAM p WITH fast : main;
  END_RESOURCE
END_CONFIGURATION

(* ---- sfcaction.st ---- *)
(* An ACTION whose body is an SFC (Ed.3 6.7.4.1; Annex A, Action : ...
   FB_Body). The chart in it evolves in the scans its action runs, the
   final scan too, and is held in the others: its steps stay, its BOOL
   action keeps its value, a step's T stands still; it is never reset
   (docs/dependencies.md). Its steps and actions are the POU's by name:
   its step i2 runs mark, an action of the outer chart.
   Outer: o0 runs sub for 20 ms, o1 waits 20 ms, and again; w0 runs
   watch every scan, after sub. In sub: i0 counts k to 2, i1 lights
   lamp and waits until i1.T is 30 ms, i2 stays.
   %QB0 the steps (o0 1, o1 2, i0 4, i1 8, i2 16), %QB1 k, %QB2 lamp,
   %QB3 how many of 10, 20, 30 ms i1.T has reached, %QB4 m.
   Worked by hand, a tick 10 ms:
   tick 0: o0, i0; cnt: k 1.                         05 01 00 00 00
   tick 1: k 2, so i0 to i1.                         09 02 00 00 00
   tick 2: cnt's final scan, k 3; lamp; i1.T 10 ms;
           o0.T 20 ms, so o0 to o1.                  09 03 01 01 00
   tick 3: sub's final scan: i1.T 20 ms.             0A 03 01 02 00
   tick 4: sub held: lamp and i1.T as they were;
           o1.T 20 ms, so o1 to o0.                  0A 03 01 02 00
   tick 5: sub again, where it was: i1.T 30 ms (the
           10 ms it was held not counted): i1 to i2. 11 03 01 03 00
   tick 6: lamp falls; i2 runs mark: m 1; o0 to o1.  11 03 00 03 01
   tick 7: sub's final scan; m 2.                    12 03 00 03 02
   reference-skip: the reference compiler takes no SFC in an action. *)
PROGRAM main
  VAR k, m : INT; lamp : BOOL; END_VAR
  VAR
    q0 AT %QB0 : USINT;
    q1 AT %QB1 : USINT;
    q2 AT %QB2 : USINT;
    q3 AT %QB3 : USINT;
    q4 AT %QB4 : USINT;
  END_VAR
  INITIAL_STEP o0 : sub(N); END_STEP
  TRANSITION FROM o0 TO o1 := o0.T >= T#20ms; END_TRANSITION
  STEP o1 : END_STEP
  TRANSITION FROM o1 TO o0 := o1.T >= T#20ms; END_TRANSITION
  INITIAL_STEP w0 : watch(N); END_STEP
  TRANSITION FROM w0 TO w0 := FALSE; END_TRANSITION
  ACTION sub :
    INITIAL_STEP i0 : cnt(N); END_STEP
    TRANSITION FROM i0 TO i1 := k >= 2; END_TRANSITION
    STEP i1 : lamp(N); END_STEP
    TRANSITION FROM i1 TO i2 := i1.T >= T#30ms; END_TRANSITION
    STEP i2 : mark(N); END_STEP
    TRANSITION FROM i2 TO i2 := FALSE; END_TRANSITION
    ACTION cnt : k := k + 1; END_ACTION
  END_ACTION
  ACTION mark : m := m + 1; END_ACTION
  ACTION watch :
    q0 := BOOL_TO_USINT(o0.X) + 2 * BOOL_TO_USINT(o1.X) + 4 * BOOL_TO_USINT(i0.X)
          + 8 * BOOL_TO_USINT(i1.X) + 16 * BOOL_TO_USINT(i2.X);
    q1 := INT_TO_USINT(k);
    q2 := BOOL_TO_USINT(lamp);
    q3 := BOOL_TO_USINT(i1.T >= T#10ms) + BOOL_TO_USINT(i1.T >= T#20ms) + BOOL_TO_USINT(i1.T >= T#30ms);
    q4 := INT_TO_USINT(m);
  END_ACTION
END_PROGRAM
CONFIGURATION c RESOURCE r ON PLC TASK t(INTERVAL := T#10ms, PRIORITY := 1); PROGRAM p WITH t : main; END_RESOURCE END_CONFIGURATION

(* ---- sfcdemo.st ---- *)
(* SFC (Ed.3 6.7; docs/behaviour/sfc.md): Prokop's demo chart. Each scan
   runs the actions, those ending first, then the transitions; an action
   runs once more after its step is left (the final scan), so the P
   action EntryCount runs twice per entry, as the standard's
   ACTION_CONTROL and CODESYS have it - P1 would run once. The reference compiler tests
   the transitions first and has no final scan: iecf's trace is
   sfcdemo.iecf.trace. *)
PROGRAM DemoSfc
VAR
    start AT %IX0.0 : BOOL;
    running AT %QX0.0 : BOOL;
    entries AT %QW1 : INT;
END_VAR

INITIAL_STEP Idle:
    IdleMode(N);
END_STEP

STEP Active:
    ActiveMode(N);
    EntryCount(P);
END_STEP

TRANSITION FROM Idle TO Active
    := start;
END_TRANSITION

TRANSITION FROM Active TO Idle
    := NOT start;
END_TRANSITION

ACTION IdleMode:
    running := FALSE;
END_ACTION

ACTION ActiveMode:
    running := TRUE;
END_ACTION

ACTION EntryCount:
    entries := entries + 1;
END_ACTION

END_PROGRAM

CONFIGURATION Config0
    RESOURCE Res0 ON PLC
        TASK task0(INTERVAL := T#10ms, PRIORITY := 0);
        PROGRAM instance0 WITH task0 : DemoSfc;
    END_RESOURCE
END_CONFIGURATION

(* ---- sfchold.st ---- *)
(* A manual mode (docs/c-output.md §3): while the platform holds the
   charts no transition is cleared, though its condition is TRUE; the
   steps stay as they are, or as the platform enters and leaves them,
   and their actions run as for any step - a P action on a step the
   platform entered, with its final scan, and the step's time from that
   entry. Freed, the chart goes on from the steps it then has. The x
   outputs show the active steps, npulse the P action's runs, late that
   S2 has been active 20 ms. A scan is 10 ms. iecf's alone (reference-skip), its
   trace checked by hand. *)
PROGRAM main
VAR
  go AT %IX0.0 : BOOL;
  x0 AT %QX0.0 : BOOL;
  x1 AT %QX0.1 : BOOL;
  x2 AT %QX0.2 : BOOL;
  npulse AT %QB1 : USINT;
  late AT %QX0.3 : BOOL;
END_VAR

INITIAL_STEP S0:
  x0(N);
END_STEP
STEP S1:
  x1(N);
END_STEP
STEP S2:
  x2(N);
  Pulse(P);
  Clock(N);
END_STEP

TRANSITION FROM S0 TO S1 := go; END_TRANSITION
TRANSITION FROM S1 TO S2 := go; END_TRANSITION
TRANSITION FROM S2 TO S0 := NOT go; END_TRANSITION

ACTION Pulse:
  npulse := npulse + 1;
END_ACTION
ACTION Clock:
  late := S2.T >= T#20ms;
END_ACTION
END_PROGRAM

CONFIGURATION c
  RESOURCE r ON cpu
    TASK t(INTERVAL := T#10ms, PRIORITY := 1);
    PROGRAM p WITH t : main;
  END_RESOURCE
END_CONFIGURATION

(* ---- sfcind.st ---- *)
(* SFC indicator variables (Ed.3 6.7.4.2, Table 58 field "c",
   deprecated; W0007): after the standard's own example, Figure 23's
   S22 to S27, in small. An indicator does nothing of its own: the
   action sets it, and a transition reads it. Actions run before the
   transitions, and a step's action once more as it is left (its final
   scan, as `sfcdemo`). Worked by hand (q0 the step whose action ran
   last, q1 the count of breaker, q2 closed):

   tick 0: S22: breaker, n 1, not closed (Q 16 01 00).
   tick 1: n 2, closed TRUE (Q 16 02 01); S22 to S23.
   tick 2: breaker's final scan, n 3, then opener resets closed (Q 17
   03 00); NOT closed: S23 to S22.
   tick 3: opener's final scan, then breaker, n 4, closed (Q 16 04 01).
   sfcind.iecf.trace: the reference compiler takes the indicator too, and
   has no final scan (as `sfcdemo`): n one less from tick 2. *)
PROGRAM main
  VAR closed : BOOL; n : USINT; st : USINT := 22; END_VAR
  VAR q AT %QB0 : USINT; q1 AT %QB1 : USINT; q2 AT %QB2 : USINT; END_VAR
  INITIAL_STEP s22 : breaker(N, closed); END_STEP
  TRANSITION FROM s22 TO s23 := closed; END_TRANSITION
  STEP s23 : opener(N); END_STEP
  TRANSITION FROM s23 TO s22 := NOT closed; END_TRANSITION
  ACTION breaker :
    st := 22;
    n := n + 1;
    closed := n >= 2;
    q := st; q1 := n; q2 := BOOL_TO_USINT(closed);
  END_ACTION
  ACTION opener :
    st := 23;
    closed := FALSE;
    q := st; q1 := n; q2 := BOOL_TO_USINT(closed);
  END_ACTION
END_PROGRAM
CONFIGURATION c RESOURCE r ON PLC TASK t(INTERVAL := T#10ms, PRIORITY := 1); PROGRAM p WITH t : main; END_RESOURCE END_CONFIGURATION

(* ---- sfcnets.st ---- *)
(* Two SFC networks in one POU (Ed.3 Annex A, SFC : Sfc_Network +),
   each with its own INITIAL_STEP, evolving side by side in each scan.
   Network A goes s0 to s1 once ca reaches 2 and straight back; network
   B goes t0 to t1 once cb reaches 3 and stays. A third, w0 alone, runs
   watch every scan: Q0 is 1 when s1 is active and 2 when t1 is (as the
   steps stand when watch runs, actions before transitions). Worked by
   hand, cnt_a and cnt_b each counting their step's scans:

   tick 0: ca 1, cb 1; s0 and t0: Q0 00.
   tick 1: ca 2, cb 2: s0's transition holds, s1 next.
   tick 2: s1 active (Q0 01); cnt_a's final scan, ca 3; cb 3: t1 next.
   tick 3: s0 again, t1 (Q0 02); cnt_b's final scan, cb 4; ca 4: s1.
   tick 4: s1 and t1 (Q0 03); cnt_a's final scan, ca 5.
   tick 5: s0 and t1 (Q0 02).
   The reference compiler's trace is the same; its ca differs (no final
   scan, as `sfcdemo`), which the trace does not show. *)
PROGRAM main
  VAR ca, cb : INT; END_VAR
  VAR q AT %QB0 : USINT; END_VAR
  INITIAL_STEP s0 : cnt_a(N); END_STEP
  TRANSITION FROM s0 TO s1 := ca >= 2; END_TRANSITION
  STEP s1 : END_STEP
  TRANSITION FROM s1 TO s0 := TRUE; END_TRANSITION
  INITIAL_STEP t0 : cnt_b(N); END_STEP
  TRANSITION FROM t0 TO t1 := cb >= 3; END_TRANSITION
  STEP t1 : END_STEP
  TRANSITION FROM t1 TO t1 := FALSE; END_TRANSITION
  INITIAL_STEP w0 : watch(N); END_STEP
  TRANSITION FROM w0 TO w0 := FALSE; END_TRANSITION
  ACTION cnt_a : ca := ca + 1; END_ACTION
  ACTION cnt_b : cb := cb + 1; END_ACTION
  ACTION watch : q := BOOL_TO_USINT(s1.X) + 2 * BOOL_TO_USINT(t1.X); END_ACTION
END_PROGRAM
CONFIGURATION c RESOURCE r ON PLC TASK t(INTERVAL := T#10ms, PRIORITY := 1); PROGRAM p WITH t : main; END_RESOURCE END_CONFIGURATION

(* ---- shadowcall.st ---- *)
(* shadowing: a call reaches the function past a local of its name that
   cannot be called, as CODESYS resolves it (found in OSCAT NETWORK's
   DLOG_CRON_TAB). Worked by hand: Twice(21) + LEN(twice) with twice the
   STRING 'x', 42 + 1 = 43 (%QW0); max := MAX(3, 7), 7 (%QW2);
   DAY_OF_WEEK(D#2026-11-19), a Thursday, 4 (%QB4).
   reference-skip: shadowing is CODESYS's, not IEC 61131-3. *)
FUNCTION Twice : INT
VAR_INPUT x : INT; END_VAR
Twice := 2 * x;
END_FUNCTION
PROGRAM main
VAR twice : STRING[10]; max : INT; d : DATE := D#2026-11-19; END_VAR
VAR q0 AT %QW0 : INT; q1 AT %QW2 : INT; q2 AT %QB4 : USINT; END_VAR
twice := 'x';
max := MAX(3, 7);
q0 := Twice(21) + LEN(twice);
q1 := max;
q2 := DAY_OF_WEEK(d);
END_PROGRAM

CONFIGURATION cf
  RESOURCE r ON x
    TASK tk(INTERVAL := T#10ms, PRIORITY := 1);
    PROGRAM p WITH tk : main;
  END_RESOURCE
END_CONFIGURATION

(* ---- single.st ---- *)
(* A TASK triggered by SINGLE, and a TASK whose INTERVAL is a variable
   (Ed.3 6.8.2: Data_Source; rules a and b). The tick is 10 ms, the
   constant task's interval.
   ev (SINGLE := %IX0.0, no INTERVAL) runs on each rising edge of
   %IX0.0, which is TRUE at ticks 1, 2, 4 and FALSE at 0, 3, 5: it runs
   at ticks 1 and 4. Its count: 0 1 1 1 2 2 (%QB0).
   both (SINGLE := go, INTERVAL := T#20ms), go a global the program c
   sets from %IX0.1, TRUE at tick 3 only (c runs first, priority 0): the
   edge at 3, and at the interval at ticks 0, 2, 4 while go is FALSE:
   it runs at 0, 2, 3, 4. Count: 1 1 2 3 4 4 (%QB1).
   per (INTERVAL := iv, iv a global the program c sets: T#20ms, then
   T#30ms from tick 3 on): at 0, 2 (20 ms), then 3 (30 ms divides 30).
   Count: 1 1 2 3 3 3 (%QB2).
   reference-skip: the reference compiler's host knows no SINGLE. *)
PROGRAM count
  VAR_INPUT go : BOOL; END_VAR
  VAR_OUTPUT n : INT; END_VAR
  n := n + 1;
END_PROGRAM
PROGRAM ctl
  VAR_EXTERNAL go : BOOL; iv : TIME; END_VAR
  VAR i1 AT %IX0.1 : BOOL; t AT %IB1 : BYTE; END_VAR
  go := i1;
  IF t >= 3 THEN
    iv := T#30ms;
  END_IF;
END_PROGRAM
PROGRAM show
  VAR_EXTERNAL a : INT; b : INT; c2 : INT; END_VAR
  VAR q0 AT %QB0 : SINT; q1 AT %QB1 : SINT; q2 AT %QB2 : SINT; END_VAR
  q0 := INT_TO_SINT(a);
  q1 := INT_TO_SINT(b);
  q2 := INT_TO_SINT(c2);
END_PROGRAM

CONFIGURATION cf
  VAR_GLOBAL go : BOOL; iv : TIME := T#20ms; a : INT; b : INT; c2 : INT; END_VAR
  RESOURCE r ON x
    TASK fast(INTERVAL := T#10ms, PRIORITY := 0);
    TASK ev(SINGLE := %IX0.0, PRIORITY := 1);
    TASK both(SINGLE := go, INTERVAL := T#20ms, PRIORITY := 2);
    TASK per(INTERVAL := iv, PRIORITY := 3);
    TASK last(INTERVAL := T#10ms, PRIORITY := 9);
    PROGRAM c WITH fast : ctl;
    PROGRAM p1 WITH ev : count(n => a);
    PROGRAM p2 WITH both : count(n => b);
    PROGRAM p3 WITH per : count(n => c2);
    PROGRAM s WITH last : show;
  END_RESOURCE
END_CONFIGURATION

(* ---- splitclamp.st ---- *)
(* A SPLIT's part stored into a subrange (Ed.3 Table 36, 6.4.4.3): the
   month 11 into a USINT (1..6) is clamped to 6 and flagged, as any store
   into a subrange (docs/dependencies.md); the day 8 into an element of an
   array of the subrange, clamped too. iecf only (reference-skip: the reference compiler has
   no SPLIT). *)
TYPE half : USINT (1..6); END_TYPE
PROGRAM main
VAR
  r_month AT %MB0 : USINT;
  r_day AT %MB1 : USINT;
  r_hour AT %MB2 : USINT;
END_VAR
VAR
  m : half := 1;
  a : ARRAY[1..2] OF half;
  h : USINT (0..23);
END_VAR
SPLIT_DT(IN := DT#2026-11-08-05:00:00, MONTH => m, DAY => a[2], HOUR => h);
r_month := m;
r_day := a[2];
r_hour := h;
END_PROGRAM

CONFIGURATION plant
  RESOURCE r ON PLC
    TASK fast(INTERVAL := T#10ms, PRIORITY := 0);
    PROGRAM p WITH fast : main;
  END_RESOURCE
END_CONFIGURATION

(* ---- splitenable.st ---- *)
(* EN and ENO on a SPLIT (Ed.3 6.6.1.5, Table 36; docs/dependencies.md).
   EN FALSE: IN is not evaluated - i is out of bounds at tick 0 and
   nothing faults - and every output keeps its value, ENO FALSE. EN TRUE:
   the parts are stored, ENO TRUE. A part that does not fit its output
   (1999 into a USINT, at tick 2) is the call's own flag: wrapped, flagged
   and ENO FALSE. iecf only (reference-skip: the reference compiler has no
   SPLIT). *)
PROGRAM main
VAR
  r_year AT %MW0 : UINT := 7;
  r_month AT %MB2 : USINT := 7;
  r_day AT %MB3 : USINT := 7;
  r_ok AT %MX4.0 : BOOL;
  r_wide AT %MX4.1 : BOOL;
  r_small AT %MB5 : USINT := 7;
END_VAR
VAR
  days : ARRAY[1..2] OF DATE := [D#2026-11-08, D#1999-12-31];
  i : INT := 3;
  run : BOOL;
  narrow : BOOL;
END_VAR
SPLIT_DATE(EN := run, IN := days[i], YEAR => r_year, MONTH => r_month, DAY => r_day, ENO => r_ok);
SPLIT_DATE(EN := narrow, IN := days[2], YEAR => r_small, ENO => r_wide);
narrow := run;
run := TRUE;
i := 1;
END_PROGRAM

CONFIGURATION plant
  RESOURCE r ON PLC
    TASK fast(INTERVAL := T#10ms, PRIORITY := 0);
    PROGRAM p WITH fast : main;
  END_RESOURCE
END_CONFIGURATION

(* ---- splitindex.st ---- *)
(* A SPLIT whose output is an array element out of bounds (Ed.3 Table 36,
   6.5.2.4): the task faults and nothing of the statement is stored - not
   the year before the bad element in the outputs' order, nor the day
   after it. At tick 0 the index is 2 and all three are stored; at tick 1
   it is 4 and the date another, and the bytes stay as tick 0 left them.
   iecf only (reference-skip: the reference compiler has no SPLIT). *)
PROGRAM main
VAR
  r_year AT %MW0 : UINT;
  r_day AT %MB2 : USINT;
  r_month AT %MB3 : USINT;
END_VAR
VAR
  i : INT := 1;
  d : DATE := D#2026-11-08;
  a : ARRAY[1..3] OF USINT;
END_VAR
i := i + 1;
SPLIT_DATE(IN := d, YEAR => r_year, MONTH => a[i], DAY => r_day);
r_month := a[2];
i := i + 1;
d := D#2027-12-09;
END_PROGRAM

CONFIGURATION plant
  RESOURCE r ON PLC
    TASK fast(INTERVAL := T#10ms, PRIORITY := 0);
    PROGRAM p WITH fast : main;
  END_RESOURCE
END_CONFIGURATION

(* ---- splitwrap.st ---- *)
(* A SPLIT's part converted to an output's type that cannot hold it
   (Ed.3 Table 36; docs/dependencies.md): the year 2026 into a USINT wraps
   to 16#EA and is flagged, as any integer conversion; the month and day
   fit. iecf only (reference-skip: the reference compiler has no SPLIT). *)
PROGRAM main
VAR
  r_year AT %MB0 : USINT;
  r_month AT %MB1 : USINT;
  r_day AT %MB2 : USINT;
END_VAR
SPLIT_DATE(D#2026-11-08, r_year, r_month, r_day);
END_PROGRAM

CONFIGURATION plant
  RESOURCE r ON PLC
    TASK fast(INTERVAL := T#10ms, PRIORITY := 0);
    PROGRAM p WITH fast : main;
  END_RESOURCE
END_CONFIGURATION

(* ---- stringchars.st ---- *)
(* One character of a STRING, s[i] (Ed.3 6.4.2), from 1, a CHAR: read,
   and written - only a character the string has: a position below 1 or
   past its end leaves s as it is, flagged STRING_POSITION; c = '$00'
   cuts the string there, as '$00' ends any string. In an array of
   strings, a[1][2], as Ed.3's Example 1; a CHAR into a STRING.
   Worked by hand, a[1] '5678' at the start: qc '6' (16#36); a[1] then
   '5668', '5666', '6666'; a[0] '6'; t 'A'.
   Tick 0, n 2: s 'AxC'.
   Tick 1, n 4: past the end, s stays 'ABC', flag STRING_POSITION on
   line 34.
   Tick 2, n 0: below 1, s stays 'ABC', still flagged.
   Tick 3, n 3: the last character, s 'ABx'; the flag stays until the
   platform clears it (docs/c-output.md).
   reference-skip: s[i] is Ed.3's; the reference compiler (Ed.2) has
   none. *)
PROGRAM main
VAR
  n AT %IB0 : SINT;
  qs AT %QB0 : STRING[4];
  qc AT %QB5 : CHAR;
  qa AT %QB6 : STRING[4];
  qz AT %QB11 : STRING[4];
  qw AT %QB16 : STRING[4];
END_VAR
VAR
  s : STRING[4];
  t : STRING[4];
  a : ARRAY[0..1] OF STRING[4] := ['1234', '5678'];
END_VAR
t := 'ABC';
t[2] := '$00';
qw := t;
s := 'ABC';
s[n] := 'x';
qs := s;
qc := a[1][2];
a[1][3] := qc;
a[1][4] := '6';
a[1][1] := a[1][4];
a[0] := a[1][4];
qa := a[1];
qz := a[0];
END_PROGRAM

CONFIGURATION Plant
  RESOURCE r ON PLC
    TASK fast(INTERVAL := T#10ms, PRIORITY := 1);
    PROGRAM p WITH fast : main;
  END_RESOURCE
END_CONFIGURATION

(* ---- strings.st ---- *)
(* STRING (Ed.3 6.4.2, Table 34): variables with and without a length,
   initial values, assignment, comparison, and LEN, LEFT, RIGHT, MID,
   CONCAT, INSERT, DELETE, REPLACE, FIND, with lengths and positions
   from the inputs, inside the strings so both compilers define them
   (the reference compiler reads no STRING[n] variable, so every one here is STRING). A
   string in a structure and in an array. The results are seen through
   LEN, FIND and comparisons. From tick 2 INSERT's P is past the end of
   its string: iecf appends and flags it (docs/dependencies.md), which
   the reference compiler does not; the bytes are the same. *)
TYPE item : STRUCT
  tag : STRING := 'ab';
  n : INT;
END_STRUCT;
END_TYPE
PROGRAM main
VAR
  l AT %IW0 : INT;
  p AT %IW2 : INT;
  r_len AT %MW0 : INT;
  r_find AT %MW2 : INT;
  r_cmp AT %MW4 : WORD;
  r_mix AT %MW6 : INT;
END_VAR
VAR
  greeting : STRING := 'hello';
  message : STRING;
  short : STRING;
  names : ARRAY[1..2] OF STRING := ['x', 'y$'z'];
  it : item;
  part : STRING;
END_VAR
message := CONCAT(greeting, ' world', '!');
r_len := LEN(message);
r_find := FIND(message, 'wor');
short := LEFT(message, 4);
part := MID(message, l, p);
r_mix := LEN(part) * 100 + FIND(message, part);
r_cmp := 0;
IF message = 'hello world!' THEN r_cmp := r_cmp OR 1; END_IF;
IF 'apple' < greeting THEN r_cmp := r_cmp OR 2; END_IF;
IF short = 'hell' THEN r_cmp := r_cmp OR 4; END_IF;
IF names[2] = 'y$'z' THEN r_cmp := r_cmp OR 8; END_IF;
it.tag := names[1];
IF it.tag <> 'x' THEN r_cmp := r_cmp OR 16; END_IF;
IF RIGHT(message, l) = 'ld!' THEN r_cmp := r_cmp OR 32; END_IF;
IF INSERT(greeting, '--', p) = 'he--llo' THEN r_cmp := r_cmp OR 64; END_IF;
IF DELETE(message, l, p) = 'hello!' THEN r_cmp := r_cmp OR 128; END_IF;
IF REPLACE(greeting, 'LL', l, p) = 'heLLo' THEN r_cmp := r_cmp OR 256; END_IF;
IF GT(message, greeting) THEN r_cmp := r_cmp OR 512; END_IF;
IF part >= 'w' THEN r_cmp := r_cmp OR 1024; END_IF;
END_PROGRAM

CONFIGURATION config
  RESOURCE res ON PLC
    TASK t(INTERVAL := T#10ms, PRIORITY := 0);
    PROGRAM p WITH t : main;
  END_RESOURCE
END_CONFIGURATION

(* ---- targetidx.st ---- *)
(* An assignment's target indexed by a FUNCTION with effects or by a
   real converted to an integer; a statement whose conversion fails is
   left undone, though its placeholder would fault.
   Inc adds 1 to its in-out and gives it. n 0. Worked by hand:
   a[Inc(n)] := 5: Inc called once, n 1, a[1] 5 (%QB0, n %QB1).
   aa[Inc(n)][Inc(n)] := 9: n 2, then 3; aa[2][3] 9 (%QB2, n %QB3).
   ps[Inc(n) - 2].x := 4: n 4, ps[2].x 4 (%QB4).
   r 2.0: a[REAL_TO_INT(r)] := 6: a[2] 6 (%QB5).
   The target first, then the value (Ed.3 7.3.2): b[Inc(n)] := n makes
   n 5, then reads it: b[5] 5 (%QB6).
   Then r is 1.0E10, beyond INT, and each statement it is converted in
   is left undone and flagged CONVERSION, first at the line of
   a[REAL_TO_INT(r)] := 7 - though the placeholder it would give, 0,
   is outside a and divides by zero: a[1] is still 5 (%QB7); v := 10 /
   REAL_TO_INT(r) leaves v 7 (%QB8); v := a[REAL_TO_INT(r)] leaves it 7
   (%QB9); IF a[REAL_TO_INT(r)] > 0 runs no branch (%QB10 stays 0).
   Last, a[i] := 1 with i 4: a fault (INDEX), nothing stored.
   reference-skip: ARRAY OF ARRAY: the reference compiler refuses it. *)
TYPE
  PT : STRUCT x : INT; END_STRUCT;
END_TYPE
FUNCTION Inc : INT
  VAR_IN_OUT io : INT; END_VAR
  io := io + 1;
  Inc := io;
END_FUNCTION
PROGRAM main
  VAR
    n : INT;
    r : REAL := 2.0;
    v : INT := 7;
    i : INT := 4;
    a : ARRAY [1..3] OF INT;
    aa : ARRAY [1..3] OF ARRAY [1..3] OF INT;
    ps : ARRAY [1..3] OF PT;
    b : ARRAY [1..9] OF INT;
  END_VAR
  VAR
    q0 AT %QB0 : SINT;
    q1 AT %QB1 : SINT;
    q2 AT %QB2 : SINT;
    q3 AT %QB3 : SINT;
    q4 AT %QB4 : SINT;
    q5 AT %QB5 : SINT;
    q6 AT %QB6 : SINT;
    q7 AT %QB7 : SINT;
    q8 AT %QB8 : SINT;
    q9 AT %QB9 : SINT;
    q10 AT %QB10 : SINT;
  END_VAR
  a[Inc(n)] := 5;
  q0 := INT_TO_SINT(a[1]);
  q1 := INT_TO_SINT(n);
  aa[Inc(n)][Inc(n)] := 9;
  q2 := INT_TO_SINT(aa[2][3]);
  q3 := INT_TO_SINT(n);
  ps[Inc(n) - 2].x := 4;
  q4 := INT_TO_SINT(ps[2].x);
  a[REAL_TO_INT(r)] := 6;
  q5 := INT_TO_SINT(a[2]);
  b[Inc(n)] := n;
  q6 := INT_TO_SINT(b[5]);
  r := 1.0E10;
  a[REAL_TO_INT(r)] := 7;
  q7 := INT_TO_SINT(a[1]);
  v := 10 / REAL_TO_INT(r);
  q8 := INT_TO_SINT(v);
  v := a[REAL_TO_INT(r)];
  q9 := INT_TO_SINT(v);
  IF a[REAL_TO_INT(r)] > 0 THEN
    q10 := 1;
  END_IF;
  a[i] := 1;
END_PROGRAM

CONFIGURATION c
  RESOURCE r ON x
    TASK t(INTERVAL := T#10ms, PRIORITY := 1);
    PROGRAM p WITH t : main;
  END_RESOURCE
END_CONFIGURATION

(* ---- tasks.st ---- *)
(* Two tasks of different intervals: which program instances run on which
   tick, in the order the configuration lists them, and two instances of
   one program, each with its own state.

   No connections to the programs' inputs and outputs: the reference compiler 7949c0b
   crashes (SIGSEGV) on a literal given to a program input,
   `counter(inc := 1)`, and the C it writes for a connection to a global
   does not compile (`B.INC = *TEN`). Ed.2 allows both. *)
PROGRAM bump
VAR
  mine : INT;
END_VAR
VAR_EXTERNAL
  total : INT;
  order : INT;
END_VAR
mine := mine + 1;
total := total + 1;
order := (order MOD 1000) * 10 + mine;
END_PROGRAM

PROGRAM report
VAR
  runs AT %MW4 : INT;
END_VAR
VAR_EXTERNAL
  total : INT;
  seen : INT;
END_VAR
runs := runs + 1;
seen := total;
END_PROGRAM

CONFIGURATION plant
  VAR_GLOBAL
    total AT %MW0 : INT;
    order AT %MW2 : INT;
    seen AT %MW6 : INT;
  END_VAR
  RESOURCE r ON PLC
    TASK fast(INTERVAL := T#10ms, PRIORITY := 1);
    TASK slow(INTERVAL := T#30ms, PRIORITY := 2);
    PROGRAM a WITH fast : bump;
    PROGRAM b WITH slow : bump;
    PROGRAM c WITH slow : report;
  END_RESOURCE
END_CONFIGURATION

(* ---- timers.st ---- *)
(* The timers of Ed.3 Table 46 against the time the platform passes in:
   TON, TOF and TP, started, held, released and restarted. ET is read in
   milliseconds with TIME arithmetic only: TIME_TO_DINT is not in Ed.3
   Figure 11. *)
FUNCTION ms : INT
VAR_INPUT
  t : TIME;
END_VAR
VAR
  i : INT;
  d : TIME;
END_VAR
ms := 0;
d := T#0ms;
FOR i := 1 TO 200 DO
  d := d + T#1ms;
  IF t >= d THEN
    ms := i;
  END_IF;
END_FOR;
END_FUNCTION

PROGRAM main
VAR
  run AT %IX0.0 : BOOL;
  pulse AT %IX0.1 : BOOL;
  on_q AT %QX0.0 : BOOL;
  off_q AT %QX0.1 : BOOL;
  tp_q AT %QX0.2 : BOOL;
  on_et AT %MW0 : INT;
  off_et AT %MW2 : INT;
  tp_et AT %MW4 : INT;
END_VAR
VAR
  t_on : TON;
  t_off : TOF;
  t_p : TP;
END_VAR
t_on(IN := run, PT := T#35ms);
t_off(IN := run, PT := T#20ms);
t_p(IN := pulse, PT := T#30ms);
on_q := t_on.Q;
off_q := t_off.Q;
tp_q := t_p.Q;
on_et := ms(t_on.ET);
off_et := ms(t_off.ET);
tp_et := ms(t_p.ET);
END_PROGRAM

CONFIGURATION plant
  RESOURCE r ON PLC
    TASK fast(INTERVAL := T#10ms, PRIORITY := 0);
    PROGRAM p WITH fast : main;
  END_RESOURCE
END_CONFIGURATION

(* ---- types.st ---- *)
(* Derived types: enumerated, subrange, ARRAY of one and two dimensions
   with bounds not at 0, STRUCT, an array of structures, initial values of
   each, and assignment of a whole structure and a whole array. *)
TYPE
  mode : (idle, filling, draining) := idle;
  percent : INT (0..100) := 50;
  point : STRUCT
    x : INT := 1;
    y : INT := -1;
  END_STRUCT;
  row : ARRAY [1..4] OF INT := [10, 20, 30, 40];
END_TYPE

PROGRAM main
VAR
  inp AT %IW0 : INT;
  r_mode AT %MB0 : BYTE;
  r_pct AT %MW2 : INT;
  r_sum AT %MW4 : INT;
  r_grid AT %MW6 : INT;
  r_pt AT %MW8 : INT;
  r_pts AT %MW10 : INT;
  r_copy AT %MW12 : INT;
END_VAR
VAR
  m : mode;
  p : percent;
  r : row;
  r2 : row;
  grid : ARRAY [-1..1, 0..2] OF INT := [1, 2, 3, 4, 5, 6, 7, 8, 9];
  pt : point;
  pt2 : point := (x := 5);
  pts : ARRAY [0..2] OF point;
  i : INT;
END_VAR
CASE m OF
  idle: IF inp > 0 THEN m := filling; END_IF;
  filling: IF inp > 10 THEN m := draining; END_IF;
  draining: IF inp <= 0 THEN m := idle; END_IF;
END_CASE;
IF m = idle THEN r_mode := 0; ELSIF m = filling THEN r_mode := 1; ELSE r_mode := 2; END_IF;
p := LIMIT(0, inp * 5, 100);
r_pct := p;
r[2] := r[2] + inp;
r_sum := 0;
FOR i := 1 TO 4 DO
  r_sum := r_sum + r[i];
END_FOR;
r_grid := grid[-1, 0] * 100 + grid[0, 1] * 10 + grid[1, 2];
pt.x := pt.x + inp;
r_pt := pt.x * 100 + pt.y + pt2.x * 10 + pt2.y;
pts[1] := pt;
pts[2].y := pts[1].x;
r_pts := pts[0].x + pts[1].x + pts[2].y;
r2 := r;
r2[1] := 0;
r_copy := r[1] + r2[1] + r2[2];
END_PROGRAM

CONFIGURATION plant
  RESOURCE r ON PLC
    TASK fast(INTERVAL := T#10ms, PRIORITY := 0);
    PROGRAM p WITH fast : main;
  END_RESOURCE
END_CONFIGURATION

(* ---- unconverted.st ---- *)
(* A REAL converted to an integer it does not fit leaves its statement
   undone and is flagged (docs/c-output.md §5, decided 2026-11-06,
   docs/dependencies.md). At tick 1, x is 1.0E10,
   beyond INT: the assignment keeps a's value, the IF and the CASE run no
   branch, the FOR does not run, the WHILE ends, the REPEAT ends after
   its first pass. At tick 2 x is back in range. The first is flagged,
   code 4 at line 29. The reference compiler's C converts out of range, which C leaves
   undefined; its trace is what x86 gives. iecf's is
   unconverted.iecf.trace. *)
PROGRAM main
VAR
  k AT %IW0 : INT;
  a AT %MW0 : INT;
  b AT %MW2 : INT;
  c AT %MW4 : INT;
  n AT %MW6 : INT;
  w AT %MW8 : INT;
  r AT %MW10 : INT;
  ticks AT %MW12 : INT;
END_VAR
VAR
  x : REAL;
  i : INT;
END_VAR
x := 100.4;
IF k >= 1 THEN
  x := 1.0E10;
END_IF;
a := REAL_TO_INT(x);
IF REAL_TO_INT(x) > 50 THEN
  b := b + 1;
ELSE
  b := b + 100;
END_IF;
CASE REAL_TO_INT(x) OF
  100: c := c + 1;
ELSE
  c := c + 100;
END_CASE;
FOR i := 1 TO REAL_TO_INT(x) / 50 DO
  n := n + 1;
END_FOR;
i := 0;
WHILE i < REAL_TO_INT(x) / 50 DO
  i := i + 1;
  w := w + 1;
END_WHILE;
i := 0;
REPEAT
  i := i + 1;
  r := r + 1;
UNTIL i >= REAL_TO_INT(x) / 50
END_REPEAT;
ticks := ticks + 1;
END_PROGRAM

CONFIGURATION plant
  RESOURCE r ON PLC
    TASK fast(INTERVAL := T#10ms, PRIORITY := 0);
    PROGRAM p WITH fast : main;
  END_RESOURCE
END_CONFIGURATION

(* ---- validbcd.st ---- *)
(* Ed.3's validate functions (6.6.2.5.15, Table 39), BCD conversions
   (6.6.2.5.2, Table 22 3a-4b, footnote d) and endianness (6.6.2.5.13,
   Table 37). Worked by hand, on a little-endian target (as the
   harness's and Prokop's are):
   MB0  IS_VALID: 1.0E38 TRUE, its tenfold (an infinity) FALSE, that minus
        itself (a NaN) FALSE, LREAL 2.5 TRUE: 2#1001, 16#09.
   MB1  IS_VALID_BCD: WORD 16#1234 TRUE, 16#12A4 FALSE, BYTE 16#99 TRUE,
        16#9A FALSE, LWORD sixteen 9s TRUE, DWORD 16#F000 FALSE: 16#15.
   MW2  WORD_BCD_TO_UINT(16#0369) = 369 (footnote d's own); MW4
        BCD_TO_INT(16#9999) = 9999; MB6 USINT_TO_BCD_BYTE(25) = 16#25
        (footnote d's); MW8 TO_BCD_WORD(UINT#1234) = 16#1234; MD10
        DWORD_BCD_TO_UDINT(16#12345678) = 12345678; ML14
        LWORD_BCD_TO_ULINT(sixteen 9s) = 9999999999999999.
   MD22 TO_BIG_ENDIAN(DWORD#16#12345678): its bytes 12 34 56 78; MW26
        TO_BIG_ENDIAN(INT#16#0102): 01 02; MB28 TO_BIG_ENDIAN(BYTE#16#12):
        not converted, 12; MD30 FROM_BIG_ENDIAN(TO_BIG_ENDIAN(16#CAFEBABE))
        is it again; MD34 TO_LITTLE_ENDIAN(16#01020304): as it is here;
        MD38 REAL 1.5 through TO_ and FROM_LITTLE_ENDIAN: 1.5; MD42 REAL
        1.5 TO_BIG_ENDIAN: its bytes 3f c0 00 00; MW46 WCHAR 'A' (16#0041)
        TO_BIG_ENDIAN, as a WORD: 00 41; MB48 TIME T#1ms TO_BIG_ENDIAN is
        16#01000000 ms, T#4h39m37s216ms: 1.
   MB50 Rec through TO_BIG_ENDIAN, packed into the image: a 11 22 33 44,
        f 01 as it is, c 01 02 03 04. MB60 Frame (relative locations)
        through TO_BIG_ENDIAN: h a1 b2, d 01 02 03 04. MB66: an
        enumerated value (bit 0) and a STRING (bit 1) as they are, Rec
        through TO_LITTLE_ENDIAN as it is here (bit 2): 2#111, 07.
   The infinity is flagged (IECF_FAULT_OVERFLOW, line 75), and stays the
   first flag; the BCD and endianness edge cases' flags are
   runtime/tests/arith.c's.
   reference-skip: the reference compiler (Ed.2) has neither IS_VALID,
   IS_VALID_BCD, BCD of a signed integer (BCD_TO_INT) nor the
   endianness functions; the BCD conversions it has are bcd.st's,
   checked against it. *)
TYPE
  Rec : STRUCT a : DWORD; f : BOOL; c : ARRAY[0..1] OF INT; END_STRUCT;
  Frame : STRUCT h AT %B0 : WORD; d AT %B2 : DINT; END_STRUCT;
  Mode : (lo, hi);
END_TYPE
PROGRAM main
VAR
  rin : Rec := (a := 16#11223344, f := TRUE, c := [16#0102, 16#0304]);
  rle : Rec;
  fin : Frame := (h := 16#A1B2, d := 16#01020304);
  m : Mode := hi;
  str : STRING := 'ab';
  big : REAL := 1.0E38;
  r1, r2, r3 : REAL;
  half : LREAL := 2.5;
  rx : REAL := 1.5;
  t : TIME;
END_VAR
VAR
  q_valid AT %MB0 : BYTE;
  q_bcd AT %MB1 : BYTE;
  u369 AT %MW2 : UINT;
  i9999 AT %MW4 : INT;
  b25 AT %MB6 : BYTE;
  w1234 AT %MW8 : WORD;
  d AT %MD10 : UDINT;
  l AT %ML14 : ULINT;
  e32 AT %MD22 : DWORD;
  e16 AT %MW26 : INT;
  e8 AT %MB28 : BYTE;
  back AT %MD30 : DWORD;
  lit AT %MD34 : DWORD;
  rr AT %MD38 : REAL;
  rb AT %MD42 : REAL;
  wc AT %MW46 : WORD;
  q_time AT %MB48 : BYTE;
  rout AT %MB50 : Rec;
  fout AT %MB60 : Frame;
  q_more AT %MB66 : BYTE;
END_VAR
r1 := big;
r2 := big * 10.0;
r3 := r2 - r2;
q_valid := 0;
IF IS_VALID(r1) THEN q_valid := q_valid OR 1; END_IF;
IF IS_VALID(r2) THEN q_valid := q_valid OR 2; END_IF;
IF IS_VALID(r3) THEN q_valid := q_valid OR 4; END_IF;
IF IS_VALID(half) THEN q_valid := q_valid OR 8; END_IF;
q_bcd := 0;
IF IS_VALID_BCD(WORD#16#1234) THEN q_bcd := q_bcd OR 1; END_IF;
IF IS_VALID_BCD(WORD#16#12A4) THEN q_bcd := q_bcd OR 2; END_IF;
IF IS_VALID_BCD(BYTE#16#99) THEN q_bcd := q_bcd OR 4; END_IF;
IF IS_VALID_BCD(BYTE#16#9A) THEN q_bcd := q_bcd OR 8; END_IF;
IF IS_VALID_BCD(LWORD#16#9999999999999999) THEN q_bcd := q_bcd OR 16; END_IF;
IF IS_VALID_BCD(DWORD#16#F000) THEN q_bcd := q_bcd OR 32; END_IF;
u369 := WORD_BCD_TO_UINT(WORD#16#0369);
i9999 := BCD_TO_INT(WORD#16#9999);
b25 := USINT_TO_BCD_BYTE(USINT#25);
w1234 := TO_BCD_WORD(UINT#1234);
d := DWORD_BCD_TO_UDINT(DWORD#16#12345678);
l := LWORD_BCD_TO_ULINT(LWORD#16#9999999999999999);
e32 := TO_BIG_ENDIAN(DWORD#16#12345678);
e16 := TO_BIG_ENDIAN(INT#16#0102);
e8 := TO_BIG_ENDIAN(BYTE#16#12);
back := FROM_BIG_ENDIAN(TO_BIG_ENDIAN(DWORD#16#CAFEBABE));
lit := TO_LITTLE_ENDIAN(DWORD#16#01020304);
rr := FROM_LITTLE_ENDIAN(TO_LITTLE_ENDIAN(rx));
rb := TO_BIG_ENDIAN(rx);
wc := WCHAR_TO_WORD(TO_BIG_ENDIAN(WCHAR#"A"));
t := TO_BIG_ENDIAN(T#1ms);
q_time := 0;
IF t = T#4h39m37s216ms THEN q_time := 1; END_IF;
rout := TO_BIG_ENDIAN(rin);
fout := TO_BIG_ENDIAN(fin);
rle := TO_LITTLE_ENDIAN(rin);
q_more := 0;
IF TO_BIG_ENDIAN(m) = hi THEN q_more := q_more OR 1; END_IF;
IF TO_BIG_ENDIAN(str) = 'ab' THEN q_more := q_more OR 2; END_IF;
IF rle.a = rin.a AND rle.c[1] = rin.c[1] THEN q_more := q_more OR 4; END_IF;
END_PROGRAM

CONFIGURATION Plant
  RESOURCE R ON PLC
    TASK fast(INTERVAL := T#10ms, PRIORITY := 1);
    PROGRAM P WITH fast : main;
  END_RESOURCE
END_CONFIGURATION

(* ---- whileranges.st ---- *)
(* WHILE loops whose guarded variable the body only steps toward the
   bound (docs/c-output.md §2, crates/iecf-codegen ranges.rs while_facts):
   their indexes proven in range and taken unchecked, the results those of
   the checked C. An insertion sort, j from i - 1 down while j >= 1; a
   search up from 1 while j <= 8, left by EXIT; a sum down from 8 while
   j > 0 by steps of 2. Eight INTs filled from %IB0 each tick:
   a[i] = (seed * (37 i + 11)) MOD 101. Worked by hand, tick 0 (seed 3):
   a = 43 53 63 73 83 93 2 12, sorted 2 12 43 53 63 73 83 93; %QW0
   a[1] * 100 + a[8] = 293 (25 01); %QW2 the first j with a[j] >= 50, 4
   (04 00); %QW4 a[8] + a[6] + a[4] + a[2] = 93 + 73 + 53 + 12 = 231
   (e7 00); %QW6 a[4], 53 (35 00). *)
PROGRAM main
VAR
  a : ARRAY[1..8] OF INT;
  i : INT; j : INT; k : INT; s : INT;
END_VAR
VAR q0 AT %QW0 : INT; q1 AT %QW2 : INT; q2 AT %QW4 : INT; q3 AT %QW6 : INT; seed AT %IB0 : BYTE; END_VAR
FOR i := 1 TO 8 DO
  a[i] := (BYTE_TO_INT(seed) * (i * 37 + 11)) MOD 101;
END_FOR;
FOR i := 2 TO 8 DO
  k := a[i];
  j := i - 1;
  WHILE j >= 1 DO
    IF a[j] <= k THEN EXIT; END_IF;
    a[j + 1] := a[j];
    j := j - 1;
  END_WHILE;
  a[j + 1] := k;
END_FOR;
q0 := a[1] * 100 + a[8];
j := 1;
WHILE j <= 8 DO
  IF a[j] >= 50 THEN EXIT; END_IF;
  j := j + 1;
END_WHILE;
q1 := j;
s := 0;
j := 8;
WHILE j > 0 DO
  s := s + a[j];
  j := j - 2;
END_WHILE;
q2 := s;
q3 := a[4];
END_PROGRAM
CONFIGURATION plant
  RESOURCE cpu ON PLC
    TASK fast(INTERVAL := T#10ms, PRIORITY := 0);
    PROGRAM p WITH fast : main;
  END_RESOURCE
END_CONFIGURATION

(* ---- wlocated.st ---- *)
(* WSTRING at an address (docs/dependencies.md): its n + 1 UTF-16 units
   back to back from its byte, each little-endian, at an odd byte too; in
   a structure and an array there, packed. Its initial value written at
   the start (not into %I); a store writes the whole string back, so
   units after its 0 stay as they were.
   Worked by hand, the input win at %IW0:
   init: qw "ab" at Q1: 61 00 62 00 00 00 00 00; qp.n 0, qp.w "z" at
   Q11: 7a 00 00 00 00 00.
   Tick 0, win 16#263A: qw := CONCAT(qw, win) "ab$263A", then qw[1] :=
   win: "$263Ab$263A" - Q1 3a 26 62 00 3a 26 00 00; qp.n := LEN(qw) 3 at
   Q9; qp.w := qw cut to "$263Ab" - Q11 3a 26 62 00 00 00; qa[1] := qp.w
   cut to "$263A" at M4: 3a 26 00 00 (qa[0] at M0 empty); q2 := qw[2] 'b'
   at Q17.
   Tick 1, win 16#0041 ('A'): CONCAT gives "$263Ab$263AA", cut to 3:
   "$263Ab$263A", qw[1] := 'A': "Ab$263A"; qp.n 3; qp.w "Ab"; qa[1] "A".
   The cuts are flagged STRING_LENGTH: first qp.w := qw in tick 0, line
   32, a flag that stays (tick 1's CONCAT cut, line 29, behind it).
   reference-skip: WCHAR and s[i] are Ed.3's. *)
TYPE pair : STRUCT n : INT; w : WSTRING[2] := "z"; END_STRUCT; END_TYPE

PROGRAM main
VAR
  win AT %IW0 : WCHAR;
  qw AT %QW1 : WSTRING[3] := "ab";
  qp AT %QW9 : pair;
  q2 AT %QW17 : WCHAR;
  qa AT %MW0 : ARRAY[0..1] OF WSTRING[1];
END_VAR
qw := CONCAT(qw, win);
qw[1] := win;
qp.n := LEN(qw);
qp.w := qw;
qa[1] := qp.w;
q2 := qw[2];
END_PROGRAM

CONFIGURATION Plant
  RESOURCE r ON PLC
    TASK fast(INTERVAL := T#10ms, PRIORITY := 1);
    PROGRAM p WITH fast : main;
  END_RESOURCE
END_CONFIGURATION

(* ---- wrefs.st ---- *)
(* REF_TO a WSTRING (Ed.3 6.4.4.10): one reference to a WSTRING at an
   address (odd byte 1, its units little-endian there) and, when pick, to
   one in C memory; what it reaches read, written whole and by s[i], and
   copied to and from; a REF_TO a structure at an address holding one.
   Worked by hand (inputs win at %IW0, pick at %IX2.0):
   tick 0, pick FALSE, win 'A' (16#41): r reaches qw "ab"; r^[1] := 'A':
   "Ab"; r^ := CONCAT(r^, '!'): "Ab!" (fits); k "Ab!"; mem := r^ "Ab!";
   qn LEN(r^) 3; rp^.w := LEFT(k, 2) "Ab", rp^.n 2; cp := rp^; qc
   cp.w[1] 'A'; qm := mem "Ab!".
   Q: 00 | qw 41 00 62 00 21 00 00 00 | qp.n 02 00 | qp.w 41 00 62 00 00
   00 | qn 03 | qc 41 00 | qm 41 00 62 00 21 00 00 00.
   Tick 1, pick TRUE, win 16#263A: r reaches mem "Ab!": "$263Ab!", then
   CONCAT "$263Ab!!" cut to "$263Ab!", flagged STRING_LENGTH at line 42,
   the first flag, which stays; mem := r^ copies it onto itself; qw
   unchanged; qp.w "$263Ab"; qc 16#263A; qm "$263Ab!".
   Tick 2, pick FALSE, win 16#E9: r reaches qw "Ab!" again: "$00E9b!";
   qp.w "$00E9b"; qc 16#E9; mem and qm "$00E9b!".
   reference-skip: WCHAR and s[i] are Ed.3's; the reference compiler
   (Ed.2) has neither. *)
TYPE pair : STRUCT n : INT; w : WSTRING[2]; END_STRUCT; END_TYPE

PROGRAM main
VAR
  win AT %IW0 : WCHAR;
  pick AT %IX2.0 : BOOL;
  qw AT %QW1 : WSTRING[3] := "ab";
  qp AT %QW9 : pair;
  qn AT %QB17 : USINT;
  qc AT %QW18 : WCHAR;
  qm AT %QW20 : WSTRING[3];
END_VAR
VAR
  mem : WSTRING[3] := "xy";
  cp : pair;
  r : REF_TO WSTRING[3];
  r2 : REF_TO WSTRING[3] := REF(mem);
  rp : REF_TO pair;
  k : WSTRING[3];
END_VAR
IF pick THEN r := REF(mem); ELSE r := REF(qw); END_IF;
r^[1] := win;
r^ := CONCAT(r^, "!");
k := r^;
r2^ := r^;
qn := INT_TO_USINT(LEN(r^));
rp := REF(qp);
rp^.w := LEFT(k, 2);
rp^.n := LEN(rp^.w);
cp := rp^;
qc := cp.w[1];
qm := mem;
END_PROGRAM

CONFIGURATION Plant
  RESOURCE r ON PLC
    TASK fast(INTERVAL := T#10ms, PRIORITY := 1);
    PROGRAM p WITH fast : main;
  END_RESOURCE
END_CONFIGURATION
